FUNCTION_BLOCK Test (* Composite Function Block Type *)
  (* Standard: 61499-2 *)
  (* Version 0.0, 7/14/2016, Andrei, nxtControl GmbH, template *)
  PACKAGE Main;
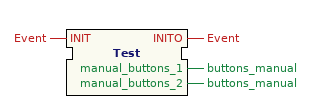
  EVENT_INPUT
    INIT; (* Initialization Request *)
  END_EVENT
  EVENT_OUTPUT
    INITO; (* Initialization Confirm *)
  END_EVENT
  PLUGS
    manual_buttons_1 : buttons_manual;
    manual_buttons_2 : buttons_manual;
  END_PLUGS
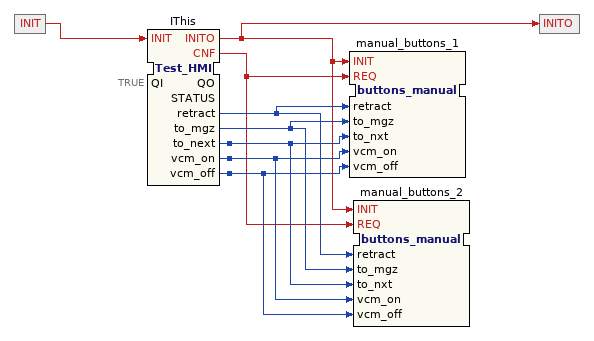
  FBS
    IThis : Test_HMI(QI := TRUE);
  END_FBS
  EVENT_CONNECTIONS
    INIT TO IThis.INIT;
    IThis.INITO TO INITO;
    IThis.INITO TO manual_buttons_1.INIT;
    IThis.INITO TO manual_buttons_2.INIT;
    IThis.CNF TO manual_buttons_1.REQ;
    IThis.CNF TO manual_buttons_2.REQ;
  END_CONNECTIONS
  DATA_CONNECTIONS
    IThis.retract TO manual_buttons_1.retract;
    IThis.retract TO manual_buttons_2.retract;
    IThis.to_mgz TO manual_buttons_1.to_mgz;
    IThis.to_mgz TO manual_buttons_2.to_mgz;
    IThis.to_next TO manual_buttons_1.to_nxt;
    IThis.to_next TO manual_buttons_2.to_nxt;
    IThis.vcm_on TO manual_buttons_1.vcm_on;
    IThis.vcm_on TO manual_buttons_2.vcm_on;
    IThis.vcm_off TO manual_buttons_1.vcm_off;
    IThis.vcm_off TO manual_buttons_2.vcm_off;
  END_CONNECTIONS
END_FUNCTION_BLOCK
